// TIA Portal V20 export
TYPE "AXIS_VIRT_N_CODE"
   STRUCT
      AXIS : Struct
         SENDING : Struct
            MC_POWER { ExternalAccessible := 'False'; ExternalVisible := 'False'; ExternalWritable := 'False'} : Struct
               ENABLE : Bool;
               START_MODE : Int;
               STOP_MODE : Int;
            END_STRUCT;
            MC_HOME { ExternalAccessible := 'False'; ExternalVisible := 'False'; ExternalWritable := 'False'} : Struct
               EXECUTE : Bool;
               POSITION : Real;
               MODE : Int;
            END_STRUCT;
            MC_MOVE_JOG { ExternalAccessible := 'False'; ExternalVisible := 'False'; ExternalWritable := 'False'} : Struct
               JOG_FORWARD : Bool;
               JOG_BACKWARD : Bool;
               VELOCITY : Real;
               POSITION_CONTROLED : Bool;
            END_STRUCT;
            MC_RESET { ExternalAccessible := 'False'; ExternalVisible := 'False'; ExternalWritable := 'False'} : Struct
               EXECUTE : Bool;
               RESTART : Bool;
            END_STRUCT;
            MC_MOVE_ABSOLUTE_JOG { ExternalAccessible := 'False'; ExternalVisible := 'False'; ExternalWritable := 'False'} : Struct
               EXECUTE : Bool;
               POSITION : Real;
               VELOCITY : Real;
               DIRECTION : Int;
            END_STRUCT;
            MC_HALT { ExternalAccessible := 'False'; ExternalVisible := 'False'; ExternalWritable := 'False'} : Struct
               EXECUTE : Bool;
            END_STRUCT;
         END_STRUCT;
         READ : Struct
            MC_POWER : Struct
               STATUS : Bool;
               BUSY : Bool;
               ERROR : Bool;
               ERROR_ID : Word;
               ERROR_INTO : Word;
            END_STRUCT;
            MC_HOME : Struct
               DONE : Bool;
               BUSY : Bool;
               COMAND_ABORTED : Bool;
               ERROR : Bool;
               ERROR_ID : Word;
               ERROR_INTO : Word;
               REFERENCE_MARK_POSITION : Real;
            END_STRUCT;
            MC_MOVE_JOG : Struct
               IN_VELOCITY : Bool;
               BUSY : Bool;
               COMAND_ABORTED : Bool;
               ERROR : Bool;
               ERROR_ID : Word;
               ERROR_INTO : Word;
            END_STRUCT;
            MC_RESET : Struct
               DONE : Bool;
               BUSY : Bool;
               ERROR : Bool;
               ERROR_ID : Word;
               ERROR_INTO : Word;
            END_STRUCT;
            MC_MOVE_ABSOLUTE : Struct
               DONE : Bool;
               BYSY : Bool;
               COMAND_ABORTED : Bool;
               ERROR : Bool;
               ERROR_ID : Word;
               ERROR_INTO : Word;
            END_STRUCT;
            MC_HALT : Struct
               done : Bool;
               BUSY : Bool;
               error : Bool;
               COMAD_ABORTED : Bool;
               ERROR_ID : Word;
               ERROR_INTO : Word;
            END_STRUCT;
         END_STRUCT;
      END_STRUCT;
   END_STRUCT;
END_TYPE
